// TIA Portal V21 export
// export: Created 2026-11-10T07:35:11.3859969Z, ExportSetting WithDefaults, DisplayName Totally Integrated Automation Portal, DisplayVersion V21 Update 3, DisplayName STEP 7 Professional, DisplayVersion V21 Update 3, DisplayName STEP 7 Safety, DisplayVersion V21, DisplayName Tech WebApplication, DisplayVersion V21, DisplayName WinCC Basic/Comfort/Advanced, DisplayVersion V21 Update 3, DisplayName WinCC Unified, DisplayVersion V21 Update 3
FUNCTION_BLOCK "FB_Lad_ex101"   // FB26, LAD
{ S7_Optimized_Access := 'TRUE' }
VERSION : 0.1
// stored: AutoNumber true, IsIECCheckEnabled false, IsRetainMemResEnabled false, MemoryReserve 100, SetENOAutomatically false, UDAEnableTagReadback false
   VAR_INPUT
      v_ob_nr : OB_ATT;
      v_event : EVENT_ATT;
      v_ret_val : Int;
   END_VAR
BEGIN

REGION Network 1: DETACH - Detach an OB from an interrupt event
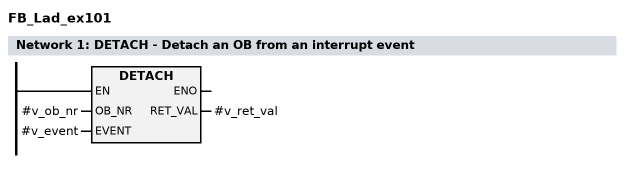
   RUNG wire#powerrail
      DETACH(OB_NR := #v_ob_nr, EVENT := #v_event, RET_VAL => #v_ret_val)
   END_RUNG
   // the same network as SCL:
   #v_ret_val := DETACH(OB_NR := #v_ob_nr, EVENT := #v_event);
END_REGION
END_FUNCTION_BLOCK
